FUNCTION_BLOCK TypeMismatch
  (* Standard: 61499-1; Description: Copyright (c) 2026 Martin Erich Jobst This program and the accompanying materials are made available under the terms of the Eclipse Public License 2.0 which is available at https://www.eclipse.org/legal/epl-2.0/ SPDX-License-Identifier: EPL-2.0 *)
  (* Version 1.0, 2026-11-18, Martin Jobst *)
  PACKAGE lib::Connection;
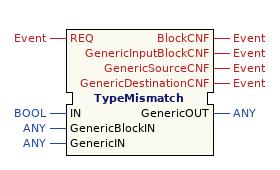
  EVENT_INPUT
    REQ;
  END_EVENT
  EVENT_OUTPUT
    BlockCNF;
    GenericInputBlockCNF;
    GenericSourceCNF;
    GenericDestinationCNF;
  END_EVENT
  VAR_INPUT
    IN : BOOL;
    GenericBlockIN : ANY;
    GenericIN : ANY;
  END_VAR
  VAR_OUTPUT
    GenericOUT : ANY;
  END_VAR
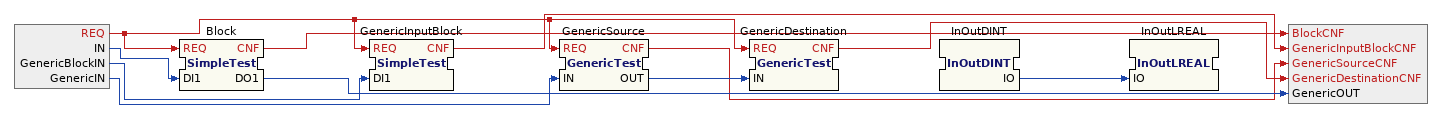
  FBS
    Block : lib::Connection::support::SimpleTest;
    GenericInputBlock : lib::Connection::support::SimpleTest;
    GenericSource : lib::Connection::support::GenericTest;
    GenericDestination : lib::Connection::support::GenericTest;
    InOutDINT : lib::Connection::support::InOutDINT;
    InOutLREAL : lib::Connection::support::InOutLREAL;
  END_FBS
  EVENT_CONNECTIONS
    REQ TO Block.REQ;
    REQ TO GenericInputBlock.REQ;
    REQ TO GenericSource.REQ;
    REQ TO GenericDestination.REQ;
    Block.CNF TO BlockCNF;
    GenericInputBlock.CNF TO GenericInputBlockCNF;
    GenericSource.CNF TO GenericSourceCNF;
    GenericDestination.CNF TO GenericDestinationCNF;
  END_CONNECTIONS
  DATA_CONNECTIONS
    IN TO Block.DI1;
    GenericBlockIN TO GenericInputBlock.DI1;
    Block.DO1 TO GenericOUT;
    GenericIN TO GenericSource.IN;
    GenericSource.OUT TO GenericDestination.IN;
    InOutDINT.IO TO InOutLREAL.IO;
  END_CONNECTIONS
END_FUNCTION_BLOCK
